(* IEC 61131-3 sources: STAR-PLC-Agent/results/raw/codex_matrix_resume_20261114/codex_deepseek/PUB003/generation/compiler_records/sim_01/precompile, 1 file *)

(* ---- FB_Task.st ---- *)
FUNCTION_BLOCK FB_Task
VAR_INPUT
    Value : REAL;
    hiLevel : REAL;
    loLevel : REAL;
    hystWindow : REAL;
END_VAR
VAR_OUTPUT
    hiAlarm : BOOL;
    loAlarm : BOOL;
    {attribute 'no_check'}
    error : BOOL;
    status : WORD;
END_VAR

error := FALSE;
status := 16#0000;

IF loLevel >= hiLevel THEN
    error := TRUE;
    status := 16#8001;
    RETURN;
END_IF

IF hystWindow >= (hiLevel - loLevel) THEN
    error := TRUE;
    status := 16#8002;
    RETURN;
END_IF

IF Value > hiLevel THEN
    hiAlarm := TRUE;
ELSIF Value < (hiLevel - hystWindow) THEN
    hiAlarm := FALSE;
END_IF

IF Value < loLevel THEN
    loAlarm := TRUE;
ELSIF Value > (loLevel + hystWindow) THEN
    loAlarm := FALSE;
END_IF
END_FUNCTION_BLOCK
